Fanuc KAREL source: KA00019.KL

PROGRAM KA00019
%NOLOCKGROUP
VAR
  SRC: REAL
  DST: XYZWPREXT
BEGIN
  SRC = 2.0
  DST = SRC
END KA00019
